{attribute 'qualified_only'}
{attribute 'strict'}
TYPE E_ValveState :
(
	Closed := 0,
	Opening,
	Open,
	Closing,
	Error := 99
);
END_TYPE

(* stored: Version 1.1.0.1
   DUT E_ValveState: Id {2ab5db84-b491-4411-a0c2-45e0010892b0} *)
